// LS Electric XG5000 project: Uas_Autoklaf
// PLC NewPLC
// module base 0 slot 0: Input/Output Module:XBM-DN32S (DC 24V INPUT/TR OUTPUT, 32points)
// module base 0 slot 1: Analog Input Module:XBF-AD04C (Volt/Current, 4-CH)
// module base 0 slot 2: Analog Output Module:XBF-DV04A (Voltage, 4-CH)

PROGRAM Autoklaf (task: Scan Program)

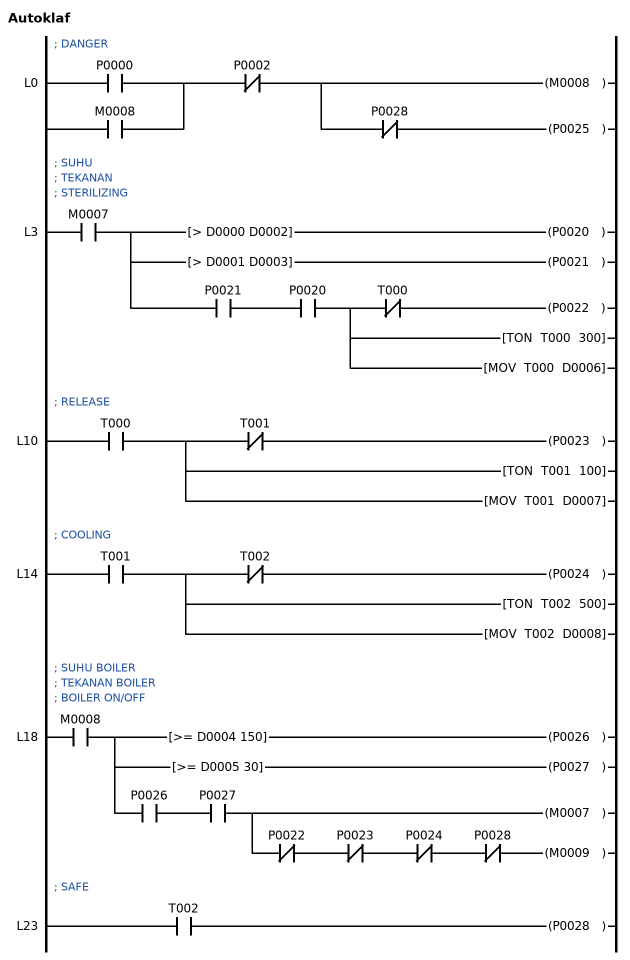
; L0
LOAD      P0000
OR        M0008
AND NOT   P0002
OUT       M0008
AND NOT   P0028
OUT       P0025
// output comment: DANGER
; L3
LOAD      M0007
MPUSH
AND>      D0000 D0002
OUT       P0020
MLOAD
AND>      D0001 D0003
OUT       P0021
MPOP
AND       P0021
AND       P0020
MPUSH
AND NOT   T000
OUT       P0022
MPOP
TON       T000 300
MOV       T000 D0006
// output comment: SUHU
// output comment: TEKANAN
// output comment: STERILIZING
; L10
LOAD      T000
MPUSH
AND NOT   T001
OUT       P0023
MPOP
TON       T001 100
MOV       T001 D0007
// output comment: RELEASE
; L14
LOAD      T001
MPUSH
AND NOT   T002
OUT       P0024
MPOP
TON       T002 500
MOV       T002 D0008
// output comment: COOLING
; L18
LOAD      M0008
MPUSH
AND>=     D0004 150
OUT       P0026
MLOAD
AND>=     D0005 30
OUT       P0027
MPOP
AND       P0026
AND       P0027
OUT       M0007
AND NOT   P0022
AND NOT   P0023
AND NOT   P0024
AND NOT   P0028
OUT       M0009
// output comment: SUHU BOILER
// output comment: TEKANAN BOILER
// output comment: BOILER ON/OFF
; L23
LOAD      T002
OUT       P0028
// output comment: SAFE